// TIA Portal V19 export
// export: Created 2026-10-15T10:10:34.9288093Z, ExportSetting WithDefaults, DisplayName Totally Integrated Automation Portal, DisplayVersion V19, DisplayName TIA Portal Openness, DisplayVersion V19, DisplayName TIA Portal Version Control Interface, DisplayVersion V19, DisplayName STEP 7 Professional, DisplayVersion V19, DisplayName STEP 7 Safety, DisplayVersion V19, DisplayName WinCC Basic/Comfort/Advanced, DisplayVersion V19, DisplayName WinCC Unified, DisplayVersion V19
FUNCTION "ROLL_TimerValue" : Word   // FC7, SCL
{ S7_Optimized_Access := 'TRUE' }
VERSION : 0.1
// stored: AutoNumber true, IsIECCheckEnabled false, SetENOAutomatically false, UDAEnableTagReadback false
   VAR_INPUT
      Number : Int;
   END_VAR
   VAR_TEMP
      count : DInt;
   END_VAR
BEGIN

   #ROLL_TimerValue := W#16#0000;
   IF (#Number < 0) OR (#Number > 127) THEN
       "ROLL_IO".ConversionFault := TRUE;
       RETURN;
   END_IF;
   IF "ROLL_State".S5Timers[#Number].BaseMs > 0 THEN
       #count := CEIL("ROLL_State".S5Timers[#Number].RemainingMs / INT_TO_LREAL("ROLL_State".S5Timers[#Number].BaseMs));
       #ROLL_TimerValue := DINT_TO_WORD(#count);
   END_IF;
END_FUNCTION
